FUNCTION_BLOCK FillValveRouter IMPLEMENTS I_FillValve, I_Cyclic
VAR
    _Name   : STRING(32);
    _Source : E_DeviceSource;
    _Chosen : I_FillValve;
END_VAR
(*
    FillValveRouter

    One I_FillValve in front of up to four candidates. The site setting,
    given once in FB_init, chooses which candidate answers and which one
    is run. A source with no candidate (0) reports a fault and is never
    open.
*)

METHOD FB_init : BOOL
VAR_INPUT
    bInitRetains    : BOOL;
    bInCopyCode     : BOOL;
    Name            : STRING(32);
    Source          : E_DeviceSource;
    FinalHardware   : I_FillValve;
    SimilarHardware : I_FillValve;
    Simulation      : I_FillValve;
    Test            : I_FillValve;
END_VAR
_Name := Name;
_Source := Source;
CASE Source OF
    E_DeviceSource.FinalHardware:   _Chosen := FinalHardware;
    E_DeviceSource.SimilarHardware: _Chosen := SimilarHardware;
    E_DeviceSource.Simulation:      _Chosen := Simulation;
    E_DeviceSource.Test:            _Chosen := Test;
END_CASE
END_METHOD

METHOD PUBLIC CyclicLogic
VAR
    Cyclic : I_Cyclic;
END_VAR
IF _Chosen <> 0 AND_THEN __QUERYINTERFACE(_Chosen, Cyclic) THEN
    Cyclic.CyclicLogic();              // only the chosen candidate runs
END_IF
END_METHOD

METHOD PUBLIC Open
IF _Chosen <> 0 THEN
    _Chosen.Open();
END_IF
END_METHOD

METHOD PUBLIC Close
IF _Chosen <> 0 THEN
    _Chosen.Close();
END_IF
END_METHOD

PROPERTY PUBLIC IsOpen : BOOL
GET
IsOpen := _Chosen <> 0 AND_THEN _Chosen.IsOpen;
END_GET
END_PROPERTY

PROPERTY PUBLIC IsClosed : BOOL
GET
IsClosed := _Chosen <> 0 AND_THEN _Chosen.IsClosed;
END_GET
END_PROPERTY

PROPERTY PUBLIC Name : STRING
GET
Name := _Name;
END_GET
END_PROPERTY

PROPERTY PUBLIC HasFault : BOOL
GET
HasFault := _Chosen = 0 OR_ELSE _Chosen.HasFault;
END_GET
END_PROPERTY

PROPERTY PUBLIC FaultText : STRING
GET
IF _Chosen = 0 THEN
    FaultText := 'No device for this source';
ELSE
    FaultText := _Chosen.FaultText;
END_IF
END_GET
END_PROPERTY

PROPERTY PUBLIC Source : E_DeviceSource
GET
Source := _Source;
END_GET
END_PROPERTY

END_FUNCTION_BLOCK

(* stored: Version 1.1.0.1, ProductVersion 3.1.4026.0
   POU FillValveRouter: Id {43b2b1bd-8c43-46e1-8f96-5f20d251f799}, SpecialFunc None
   Folder I_FillValve: Id {78a38160-681e-41d0-ac09-f902fd60cfb1}
   Folder I_Diagnosable: Id {5ba4f0b3-65eb-49e7-b7f9-e198beffb35b}
   Folder I_Cyclic: Id {a40dad8e-c43b-4a19-9a43-9595b3a05ecc}
   Method FB_init: Id {3898d12b-dd24-4801-ba44-53591b5dda70}
   Method CyclicLogic: Id {db5e4f5d-90fd-494f-bbd1-38b4ec530226}
   Method Open: Id {3bd6bfd4-1210-47d3-aade-8d140afd5d8d}
   Method Close: Id {fbd055d6-8b76-4759-86fa-50c9eb554f57}
   Property IsOpen: Id {3147a70b-f2dd-4c39-ad64-b12222a632e5}
   Get Get: Id {06b6970a-fc73-484d-af25-f8bc34371284}
   Property IsClosed: Id {47674bd4-68c3-4600-8e32-a84d8942dd1a}
   Get Get: Id {94d63ad2-9caa-43df-b9fc-c6dbecd98dc0}
   Property Name: Id {7853ee77-e746-4f5d-990b-6700e4676038}
   Get Get: Id {b477168a-597b-4172-b002-9129e3e094fe}
   Property HasFault: Id {7128146a-2abd-42b5-8b18-7c2f9560e5ca}
   Get Get: Id {049ddcdc-bae0-4c32-832d-aef2d608b0a0}
   Property FaultText: Id {892597db-190d-4fd9-aa85-3cb9c0a324a6}
   Get Get: Id {d33a5729-3129-46a7-884f-343ba138382a}
   Property Source: Id {7fc3c4be-5eb2-4b40-b216-c59fadaf26b1}
   Get Get: Id {7399d212-b68a-4cc5-a2c8-ed526745dfa1} *)
